TYPE ST_EncoderData :
STRUCT
    //------------------------------------------------------------------
    // Inputs — from EL5112 PDOs
    //------------------------------------------------------------------
    nStatusWord         : WORD;
    bInputA             : BOOL;
    bInputB             : BOOL;
    bInputC             : BOOL;
    bCounterUnderflow   : BOOL;
    bCounterOverflow    : BOOL;
    bLatchValid         : BOOL;
    bError              : BOOL;
    nCounterValue       : DWORD;
    nFrequencyValue     : DWORD;
    nState              : BYTE;
    fPosition           : LREAL;    // Scaled position [engineering units]

    //------------------------------------------------------------------
    // Outputs — written to EL5112 PDOs
    //------------------------------------------------------------------
    nSetCounterValue    : DWORD;    // Value to write to counter
    bSetCounter         : BOOL;     // Rising edge = write nSetCounterValue
    bZeroPosition       : BOOL;     // Rising edge = set counter to 0
END_STRUCT
END_TYPE

(* stored: Version 1.1.0.1, ProductVersion 3.1.4026.18
   DUT ST_EncoderData: Id {3d83a2be-9bb1-4433-8573-0e41ecf6b20e} *)
